Fanuc KAREL source: KD00018.KL

PROGRAM KD00018
%NOLOCKGROUP
VAR
  I: INTEGER
  J: INTEGER
  B: BOOLEAN
  R: REAL
  S: STRING[80]
BEGIN
  SIGNAL EVENT[1]
END KD00018
